(* IEC 61131-3 sources: codesys-build/examples/frame-assembly/src/generated/types/ST_LineDiverter, 3 files *)

(* ---- ST_LineDiverter.st ---- *)
(*
Card controls, routing context, and transfer status for an Intelligrated diverter assembly with two CS1001 cards, a ZoneMax device, and approximately two or three B&R X67 modules.
https://www.scribd.com/document/823553754/MDR-710-With-WWL-Installation-and-Maintenance-Manual
*)
TYPE ST_LineDiverter :
STRUCT
	(* Two Intelligrated CS1001 cards in the diverter assembly; each card has its own control outputs and feedback. *)
	Cards : ARRAY[1..2] OF ST_LineCS1001;
	(* Transfer sequence observations; these are not CS1001 registers. *)
	Status : ST_LineDiverterStatus;
	(* PLC-owned routing context, never mapped directly to electrical outputs. *)
	Routing : ST_LineDiverterRouting;
END_STRUCT
END_TYPE

(* ---- ST_LineDiverterRouting.st ---- *)
(*
Card controls, routing context, and transfer status for an Intelligrated diverter assembly with two CS1001 cards, a ZoneMax device, and approximately two or three B&R X67 modules.
https://www.scribd.com/document/823553754/MDR-710-With-WWL-Installation-and-Maintenance-Manual
*)
TYPE ST_LineDiverterRouting :
STRUCT
	(* 0=unknown; 1..4=configured carrier lane. Unknown must hold. *)
	CarrierDestination : INT;
	(* Identity to which the requested route applies. *)
	CommandPayload : STRING(80);
	(* LineConstants.Destination*: 0=unknown, 1=framing, 2=canvas, 3=oversize. *)
	DestinationType : INT;
	(* Payload is a bin with no remaining orders. *)
	EmptyBin : BOOL;
	(* Payload contains work requiring QC intervention. *)
	HasQC : BOOL;
	(* Derived from receiving sensors, enable state, and reservations; not a scanner observation. *)
	ReceivingAvailable : BOOL;
	(* Assigned station identity. Direction is resolved by configured port mapping. *)
	TargetStation : STRING(80);
END_STRUCT
END_TYPE

(* ---- ST_LineDiverterStatus.st ---- *)
(*
Card controls, routing context, and transfer status for an Intelligrated diverter assembly with two CS1001 cards, a ZoneMax device, and approximately two or three B&R X67 modules.
https://www.scribd.com/document/823553754/MDR-710-With-WWL-Installation-and-Maintenance-Manual
*)
TYPE ST_LineDiverterStatus :
STRUCT
	(* FALSE until the owning PLC logic supplies a current status; FALSE on stale or unavailable inputs. *)
	Valid : BOOL;
	(* Committed transfer route, not a measured actuator position. LineConstants.Route*: 0=none/hold, 1=through, 2=left, 3=right. Logical ports; no actuator wiring implied. *)
	ActiveRoute : INT;
	(* Transfer is in progress until configured arrival feedback completes it. *)
	Busy : BOOL;
	(* Fault in the actuator interface or transfer sequence. *)
	Faulted : BOOL;
	(* Payload currently committed to a transfer; cleared once arrival is confirmed. *)
	TransferPayload : STRING(80);
END_STRUCT
END_TYPE
